GLOBALCONSTANTS Etp (* Konstanten für Übungen 149-149d (ETP zwischen zwei logiBUS) *)
  (* Standard: 61499-1; Description: Copyright (c) 2026 Meisterschulen am Ostbahnhof This program and the accompanying materials are made available under the terms of the Eclipse Public License 2.0 which is available at https://www.eclipse.org/legal/epl-2.0/ SPDX-License-Identifier: EPL-2.0 *)
  (* Version 1.0, 2026-11-17, Franz Höpfinger, Meisterschulen am Ostbahnhof, ETP Partner-Filter *)
  PACKAGE Uebungen::const::Uebung_140_149;
  IMPORT isobus::pgn::NAMEFIELD_T;
  VAR_GLOBAL CONSTANT
    LOGIBUS_ADD : isobus::pgn::NAMEFIELD_T := (bSelfConf := TRUE, bIndGroup := 2, bDevClassInst := 0, bDevClass := 0, bReserved := FALSE, bFunction := 128, bFunctionInst := 0, bEcuInstance := 0, wManufCode := 1116, dwIdentNumb := 0); (* logiBUS CAN1: Hersteller 1116, Funktion 128 *)
    LOGIBUS_FLT : isobus::pgn::NAMEFIELD_T := (bSelfConf := FALSE, bIndGroup := 0, bDevClassInst := 0, bDevClass := 0, bReserved := FALSE, bFunction := 16#FF, bFunctionInst := 0, bEcuInstance := 0, wManufCode := 16#7FF, dwIdentNumb := 0); (* prüft nur wManufCode und bFunction *)
  END_VAR
END_GLOBALCONSTANTS
